FUNCTION_BLOCK FB_OverrideSelection_1
(*

The function block used to select override of axis.

Constructor: 		Patryk Panylo
Company:		E. Riexinger GmbH
Date:			23.04.2015
Version:			1.00

Date:			Revision:		Who:				Comment
dd.mm.yyyy		x.xx			Initials			comment

*)
VAR_INPUT
	(* Input variables / Eingang Variablen *)
	bEnable						:BOOL;						(* Signal FB enable *)
	rGlobalOverride				:REAL;						(* Global override *)
	rAcc							:REAL;						(* Accerlation of Override [%/s] *)
	rDec						:REAL;						(* Decerlation of Override [%/s] *)
END_VAR
VAR_OUTPUT
	(* Output variables / Ausgang Variablen *)
	rActOverride					:REAL;						(* Actual override *)
	bActGlobalOverride			:BOOL;						(* Actual override is global *)
	bActLocalOverride			:BOOL;						(* Actual override is local *)
END_VAR
VAR_IN_OUT
	(* Input Output variables / Ausgang Variablen *)
	rLocalOverride				:REAL;						(* Actual override *)
END_VAR
VAR
	(* Enummerations *)

	(* Variables *)
	rCacheGlobalOverride			:REAL;						(* Caches global override *)
	rCacheLocalOverride			:REAL;						(* Caches local override *)

	bFirstTime					:BOOL;						(* First run *)

	(* References *)

	(* Interfaces *)

	(* Instances *)
	tonChkCycleTime				:TON;						(* Check cycle time *)
END_VAR
VAR CONSTANT

END_VAR


IF NOT bEnable
THEN
	bFirstTime := FALSE;                               		(* Firstrun *)
	rActOverride := 0.0;                               		(* Override to set *)
	bActGlobalOverride := FALSE;                       	(* Actual override is global *)
	bActLocalOverride := FALSE;                       	(* Actual override is local *)
	RETURN;
END_IF;

IF NOT bFirstTime
THEN
	rCacheGlobalOverride := rGlobalOverride;          	(* Cache values *)
	rCacheLocalOverride := rLocalOverride;            		(* Cache values *)
	bActGlobalOverride := TRUE;                        			(* Actual override is global *)
	bActLocalOverride := FALSE;                       			(* Actual override is local *)
	bFirstTime := TRUE;                                				(* Firstrun *)
END_IF;

A_SelectLocal();
A_SelectGlobal();

ACTION A_SelectGlobal:

IF rCacheGlobalOverride <> rGlobalOverride
    OR rLocalOverride >= rGlobalOverride
THEN
	rCacheGlobalOverride := rGlobalOverride;
	rActOverride := rGlobalOverride;
	bActGlobalOverride := TRUE;                       	 		(* Actual override is global *)
	bActLocalOverride := FALSE;                        			(* Actual override is local *)
	rLocalOverride := rGlobalOverride;                		(* Set local Override *)
	rCacheLocalOverride := rGlobalOverride;           		(* Set local Override *)
END_IF;
END_ACTION

ACTION A_SelectLocal:

IF rCacheLocalOverride <> rLocalOverride
    AND rLocalOverride < rGlobalOverride
THEN
	rCacheLocalOverride := rLocalOverride;
	rActOverride := rLocalOverride;
	bActGlobalOverride := FALSE;                       			(* Actual override is global *)
	bActLocalOverride := TRUE;                        			(* Actual override is local *)
END_IF;
END_ACTION

END_FUNCTION_BLOCK

(* stored: Version 1.1.0.1, ProductVersion 3.1.4024.15
   POU FB_OverrideSelection_1: Id {c383340f-5b1e-4b2c-a722-a7c4273b4050}, SpecialFunc None
   Action A_SelectGlobal: Id {0bb83f9b-6914-409e-a239-5bfbd28ec4c5}
   Action A_SelectLocal: Id {2e08b69b-95e7-4b47-9a34-85eec6184436} *)
